// TIA Portal V19 export
TYPE "EM03_Input"
   STRUCT
      Cmds { S7_SetPoint := 'True'} : "EM_Input";   // Comandos estÃ¡ndar de la unidad (Start, Stop, Hold, Reset, Auto, etc.)
      CtrlMode : Int;   // 0=Off, 1=Local PID, 2=External PID (SeedMaster), 3=Water Injection
      SelectedValveIndex : Int;   // Ãndice de la vÃ¡lvula On/Off a activar (1..N)
      OpenThreshold : Real := 5.0;   // Umbral % de apertura de la vÃ¡lvula proporcional para abrir la On/Off
      CloseThreshold : Real := 3.0;   // Umbral % de apertura de la vÃ¡lvula proporcional para cerrar la On/Off
      FeedSP : Real;   // Setpoint de nivel del tacho para modo local
      WashSP : Real;   // Setpoint de nivel del tacho para lavado
      MinLevelPermit : Bool;   // Interbloqueo de nivel mÃ­nimo en tacho (LT-112)
      FeedSMMV : Real;   // Variable manipulada enviada desde SeedMaster (0..100%)
      WashMode : Bool;   // CtrlMode 3: TRUE=Lavado, FALSE=Pausa (agua segÃºn PidL)
      StableBand : Real := 2.0;   // Banda de estabilizaciÃ³n alrededor del SP (unidades de PV)
      StableTime : Time := T#10S;   // Tiempo dentro de banda para declarar COMPLETED
   END_STRUCT;
END_TYPE
